// TIA Portal V20 export
// export: Created 2026-10-20T12:50:54.8389254Z, ExportSetting WithDefaults, DisplayName Totally Integrated Automation Portal, DisplayVersion V20 Update 6, DisplayName TIA Portal Openness, DisplayVersion V20 Update 6, DisplayName TIA Portal Version Control Interface, DisplayVersion V20 Update 6, DisplayName SINAMICS Startdrive Advanced, DisplayVersion V20 SP1, DisplayName SINAMICS Startdrive G130, G150, S120, S150, SINAMICS MV, G220, S200, S210, DisplayVersion V20 SP1, DisplayName SINAMICS Startdrive G110M, G120, G120C, G120D, G120P, G115D, DisplayVersion V20 SP1, DisplayName STEP 7 Professional, DisplayVersion V20 Update 6, DisplayName STEP 7 Safety, DisplayVersion V20 Update 2, DisplayName WinCC Basic/Comfort/Advanced, DisplayVersion V20 Update 6, DisplayName WinCC Unified, DisplayVersion V20 Update 6
FUNCTION "HMI_SAFETY_FC" : Void   // FC43, F_FBD
{ S7_Optimized_Access := 'TRUE' }
VERSION : 0.1
// stored: AutoNumber true, IsIECCheckEnabled false, UDAEnableTagReadback false
   VAR_INPUT
      HMI_Box_Connected : Int;
      HMI_Reset : Bool;
      HMI_EStop : Bool;
      HMI_Profinet_Error : Bool;
      Local_Mode : Bool;
   END_VAR
   VAR_OUTPUT
      HMI_Estop_Pressed_1 : Bool;
      HMI_Estop_Pressed_2 : Bool;
      HMI_Estop_Pressed_3 : Bool;
      HMI_Estop_Pressed_4 : Bool;
      HMI_Estop_Pressed_5 : Bool;
      Reset_Comissioning_1 : Bool;
      Reset_Comissioning_2 : Bool;
      Reset_Comissioning_3 : Bool;
      Reset_Comissioning_4 : Bool;
      Reset_Comissioning_5 : Bool;
   END_VAR
   VAR_TEMP   // added for the SCL form of the ladder/FBD networks
      _w1 : Bool;
   END_VAR
BEGIN

REGION Network 1: HMI CONNECTED IN THE SYSTEM 1
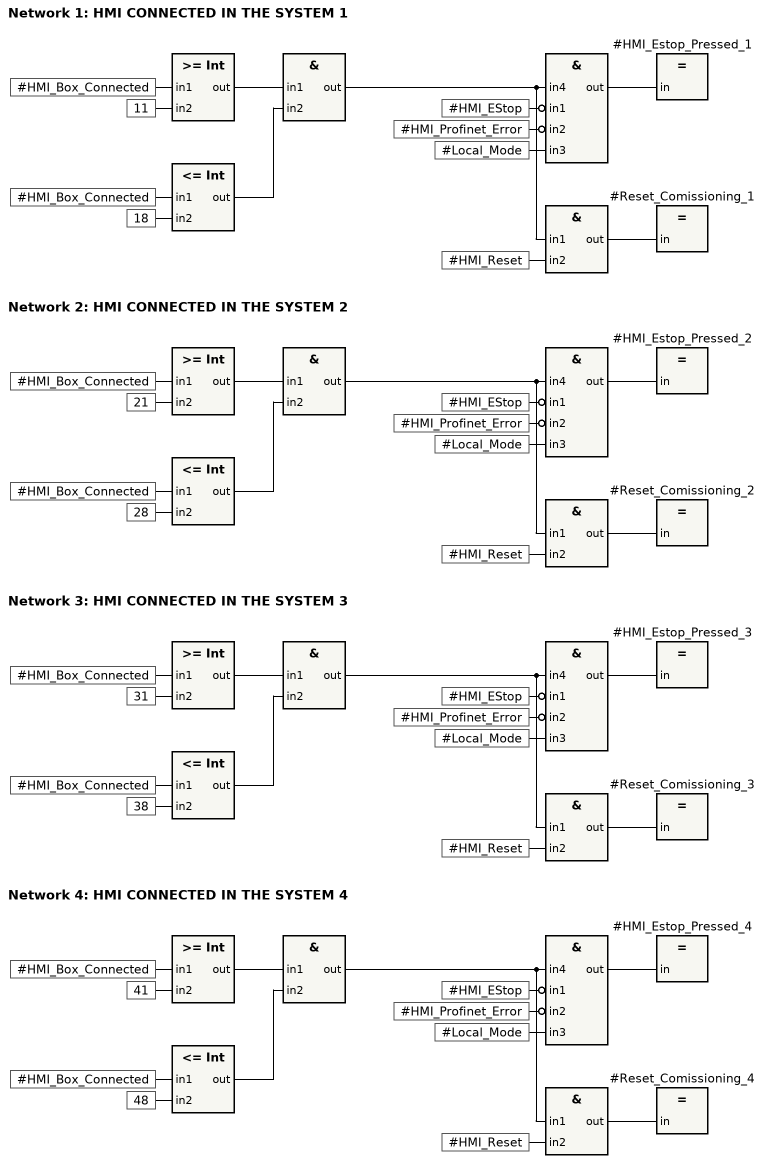
   #_w1 := (#HMI_Box_Connected >= 11) AND (#HMI_Box_Connected <= 18);
   #HMI_Estop_Pressed_1 := #_w1 AND NOT #HMI_EStop AND NOT #HMI_Profinet_Error AND #Local_Mode;
   #Reset_Comissioning_1 := #_w1 AND #HMI_Reset;
END_REGION

REGION Network 2: HMI CONNECTED IN THE SYSTEM 2
   #_w1 := (#HMI_Box_Connected >= 21) AND (#HMI_Box_Connected <= 28);
   #HMI_Estop_Pressed_2 := #_w1 AND NOT #HMI_EStop AND NOT #HMI_Profinet_Error AND #Local_Mode;
   #Reset_Comissioning_2 := #_w1 AND #HMI_Reset;
END_REGION

REGION Network 3: HMI CONNECTED IN THE SYSTEM 3
   #_w1 := (#HMI_Box_Connected >= 31) AND (#HMI_Box_Connected <= 38);
   #HMI_Estop_Pressed_3 := #_w1 AND NOT #HMI_EStop AND NOT #HMI_Profinet_Error AND #Local_Mode;
   #Reset_Comissioning_3 := #_w1 AND #HMI_Reset;
END_REGION

REGION Network 4: HMI CONNECTED IN THE SYSTEM 4
   #_w1 := (#HMI_Box_Connected >= 41) AND (#HMI_Box_Connected <= 48);
   #HMI_Estop_Pressed_4 := #_w1 AND NOT #HMI_EStop AND NOT #HMI_Profinet_Error AND #Local_Mode;
   #Reset_Comissioning_4 := #_w1 AND #HMI_Reset;
END_REGION

REGION Network 5: HMI CONNECTED IN THE SYSTEM 5
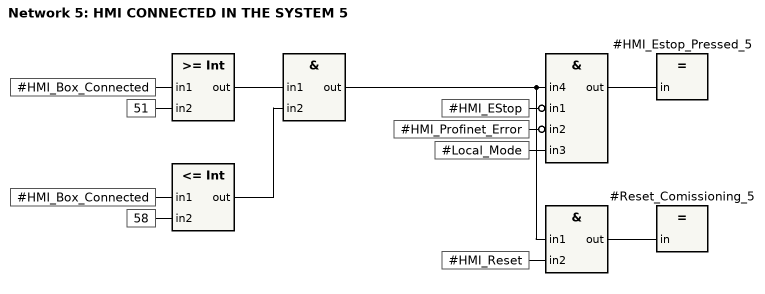
   #_w1 := (#HMI_Box_Connected >= 51) AND (#HMI_Box_Connected <= 58);
   #HMI_Estop_Pressed_5 := #_w1 AND NOT #HMI_EStop AND NOT #HMI_Profinet_Error AND #Local_Mode;
   #Reset_Comissioning_5 := #_w1 AND #HMI_Reset;
END_REGION
END_FUNCTION
